Universal Robots URScript: Feature.script

def Feature():
  # Default parameters:
  global speed_ms = 0.3
  global speed_rads = 0.75
  global accel_mss = 3
  global accel_radss = 1.2
  global blend_radius_m = 0.001

  # Add subprograms here
  # Subprogram SubProg
  def SubProg():
    # Inside sub
  end

  # Subprogram Spaced Name
  def Spaced Name():
    # Spaced body
  end

  # Subprogram Long_Program Name12
  def Long_Program Name12():
    # Long body
    set_tcp(p[0.010000, 0.000000, 0.150000, 0.000000, 0.000000, 0.000000])
    movel([-4.170995, -1.248690, 4.822082, -2.397933, 1.001165, -2.483057],accel_mss,speed_ms,0,blend_radius_m)
  end

  # Subprogram ThreadProg
  def ThreadProg():
    # Thread body
  end

  # Start of main program
  # Program generated by RoboDK v5.9.4 for UR10 on 26/10/2026 01:01:20
  # Using nominal kinematics.
  # set_reference(p[0.036764, 0.400000, 0.728939, 0.000000, 0.000000, 30.000000])
  set_tcp(p[0.000000, 0.000000, 0.120000, 0.000000, 15.000000, 0.000000])
  movej([-4.065387, -1.176966, 4.792364, -2.498712, 1.044735, -2.370328],accel_radss,speed_rads,0,blend_radius_m)
  speed_ms = 0.250
  blend_radius_m = 0.005
  movej([-4.065387, -1.176966, 4.792364, -2.498712, 1.044735, -2.370328],accel_radss,speed_rads,0,blend_radius_m)
  movel([-4.169178, -1.189198, 4.787147, -2.423562, 1.001865, -2.481067],accel_mss,speed_ms,0,blend_radius_m)
  movel([-4.113759, -1.156567, 4.786157, -2.486893, 1.024078, -2.421216],accel_mss,speed_ms,0,blend_radius_m)
  movec([-4.170995, -1.248690, 4.822082, -2.397933, 1.001165, -2.483057],[-4.077161, -1.244473, 4.849644, -2.482296, 1.039602, -2.382599],accel_mss,speed_ms,blend_radius_m)
  blend_radius_m = -0.001
  speed_rads = 0.785
  accel_mss = 0.800
  speed_ms = 0.120
  movel([-4.065387, -1.176966, 4.792364, -2.498712, 1.044735, -2.370328],accel_mss,speed_ms,0,blend_radius_m)
  movel([-4.100282, -1.212643, 4.823761, -2.538190, 1.101200, -2.039294],accel_mss,speed_ms,0,blend_radius_m)
  movej([-4.065387, -1.176966, 4.792364, -2.498712, 1.044735, -2.370328],accel_radss,speed_rads,0,blend_radius_m)
  accel_radss = 3.491
  speed_rads = 1.047
  accel_mss = 1.500
  speed_ms = 0.300
  accel_radss = 2.618
  accel_mss = 0.050
  set_standard_digital_out(5, True)
  set_standard_digital_out(3, False)
  while (get_standard_digital_in(2) != True):
    sync()
  end
  while (get_standard_digital_in(4) != False):
    sync()
  end
  sleep(1.5000)
  popup("Paused. Press continue to continue.","Message",False,False)
  sleep(2)
  # A comment line
  popup("A message","Message",False,False)
  SubProg()
  SpacedName()
  ExternalProg()
  Long_ProgramName12()
  AnotherLong_ExternalName()
  SetRPM700
  Ab_c()
  custom_code(1)
  run ThreadProg()
  set_standard_digital_out(2, 3.5)
  # set_reference(p[0.076764, 0.370000, 0.748939, 0.000000, 0.000000, 0.000000])
  set_tcp(p[0.010000, 0.000000, 0.150000, 0.000000, 0.000000, 0.000000])
  movej([-3.881380, -1.040489, 4.605461, -2.234475, 0.927523, -2.753769],accel_radss,speed_rads,0,blend_radius_m)
  movej([-4.065387, -1.176966, 4.792364, -2.498712, 1.044735, -2.370328],accel_radss,speed_rads,0,blend_radius_m)
  movel([-3.857462, -1.053266, 4.649728, -2.283236, 0.933416, -2.724861],accel_mss,speed_ms,0,blend_radius_m)
  set_tcp(p[0.000000, 0.000000, 0.120000, 0.000000, 15.000000, 0.000000])
  # set_reference(p[0.036764, 0.400000, 0.728939, 0.000000, 0.000000, 30.000000])
  movej([-4.065387, -1.176966, 4.792364, -2.498712, 1.044735, -2.370328],accel_radss,speed_rads,0,blend_radius_m)
  # End of main program
end

Feature()
